{attribute 'qualified_only'}
{attribute 'strict'}
{attribute 'to_string'}
TYPE E_Sparse :
(
	eOptionA := -10,
	eOptionB := 0,
	eOptionC := 100
);
END_TYPE

(* stored: Version 1.1.0.1, ProductVersion 3.1.4026.19
   DUT E_Sparse: Id {ddd30cc9-69f6-42a6-90c4-2cb169ac3acd} *)
